(* IEC 61131-3 sources: axsharp/src/ix.compiler/src/Ix.ixc-doc/samples/ax/src, 10 files *)

(* ---- measurement.st ---- *)
NAMESPACE MeasurementExample
    {#ix-attr:[Container(Layout.Wrap)]}
    {#ix-attr:[Group(GroupLayout.GroupBox)]}
    CLASS PUBLIC Measurement
        VAR PUBLIC
            {#ix-set:AttributeName = "Minimum"}
            Min : REAL;
            {#ix-set:AttributeName = "Measured"}
            {#ix-attr:[ReadOnly()]}
            Acquired : REAL;
            {#ix-set:AttributeName = "Maximum"}
            Max : REAL;
            {#ix-set:AttributeName = "Measurement Result"}
            Result : Result;
        END_VAR
    END_CLASS

    TYPE
        Result : INT (
            None := 0,
            Passed := 10,
            Failed := 20
        );
    END_TYPE

    CLASS PUBLIC Measurements
        VAR PUBLIC
            {#ix-attr:[Container(Layout.Stack)]}
            {#ix-attr:[Group(GroupLayout.GroupBox)]}
            {#ix-set:AttributeName = "Stack panel"}
            measurement_stack : Measurement;

            {#ix-attr:[Container(Layout.Wrap)]}
            {#ix-attr:[Group(GroupLayout.GroupBox)]}
            {#ix-set:AttributeName = "Wrap panel"}
            measurement_wrap : Measurement;

            {#ix-attr:[Container(Layout.UniformGrid)]}
            {#ix-attr:[Group(GroupLayout.GroupBox)]}
            {#ix-set:AttributeName = "Grid"}
            measurement_grid : Measurement;

            {#ix-attr:[Container(Layout.Tabs)]}
            {#ix-attr:[Group(GroupLayout.GroupBox)]}
            {#ix-set:AttributeName = "Tabs"}
            measurement_tabs : Measurement;
        END_VAR
    END_CLASS
END_NAMESPACE

(* ---- weather.st ---- *)
{#ix[Container(Layout.Tabs)]}
CLASS weather
    VAR PUBLIC
        GeoLocation : GeoLocation;
        {#ix[Container(Layout.Wrap)]}
        Temperature : REAL;
        Humidity : REAL;
        Location : STRING;
        ChillFactor : REAL;
        Feeling : Feeling;
    END_VAR
END_CLASS

CLASS weathers
    VAR PUBLIC
        i : ARRAY[0..50] OF weatherBase;
    END_VAR
END_CLASS

TYPE
    Feeling : (Freezing, Cold, Lookworm, Warm, Hot);
END_TYPE

TYPE
    Colors : INT (
        RED := 12,
        GREEN := 14,
        BLUE := 23
    );
END_TYPE

(* ---- all_primitives.st ---- *)
CLASS all_primitives
    VAR PUBLIC
        myBOOL	        :       BOOL	      ;
        myBYTE	        :       BYTE	      ;
        myWORD	        :       WORD	      ;
        myDWORD	        :       DWORD	      ;
        myLWORD	        :       LWORD	      ;
        mySINT	        :       SINT	      ;
        myINT	        :       INT	          ;
        myDINT	        :       DINT	      ;
        myLINT	        :       LINT	      ;
        myUSINT	        :       USINT	      ;
        myUINT	        :       UINT	      ;
        myUDINT	        :       UDINT	      ;
        myULINT	        :       ULINT	      ;
        myREAL	        :       REAL	      ;
        myLREAL	        :       LREAL	      ;
        myTIME	        :       TIME	      ;
        myLTIME	        :       LTIME	      ;
        myDATE	        :       DATE	      ;
     //   myLDATE	        :       LDATE	      ;
        myTIME_OF_DAY	:       TIME_OF_DAY	  ;
     //   myLTIME_OF_DAY	:       LTIME_OF_DAY  ;
        myDATE_AND_TIME  :      DATE_AND_TIME ;
     //   myLDATE_AND_TIME :      LDATE_AND_TIME;
     //   myCHAR	        :       CHAR	      ;
     //   myWCHAR	        :       WCHAR	      ;
        mySTRING	        :   STRING	      ;
        myWSTRING	    :       WSTRING	      ;
    END_VAR

END_CLASS

(* ---- example.st ---- *)
CLASS example
    VAR PUBLIC
        {#ix-attr:[Container(Layout.Stack)]}
        primitives_stack: test_primitive;
        {#ix-attr:[Container(Layout.Wrap)]}
        primitives_wrap: test_primitive;
        {#ix-attr:[Container(Layout.Tabs)]}
        primitives_tabs: test_primitive;
        {#ix-attr:[Container(Layout.UniformGrid)]}
        primitives_uniform: test_primitive;

        {#ix-attr:[Container(Layout.Stack)]}
        {#ix-attr:[Group(GroupLayout.GroupBox)]}
        test_groupbox: test_primitive;

        {#ix-attr:[Container(Layout.Stack)]}
        {#ix-attr:[Group(GroupLayout.Border)]}
        test_border: test_primitive;

        {#ix-attr:[Container(Layout.Tabs)]}
        {#ix-attr:[Group(GroupLayout.GroupBox)]}
        testgroupbox: groupbox;
        testborder: border;

        ixcomponent_instance: ixcomponent;
        ixcomponent_instance2: MySecondNamespace.ixcomponent;
        ixcomponent_instance3: ThirdNamespace.ixcomponent;

        refIxComponent : REF_TO ixcomponent;
    END_VAR

    METHOD PUBLIC ReferenceToComponent : Int
        refIxComponent^ := ixcomponent_instance;
    END_METHOD

END_CLASS

(* ---- geolocation.st ---- *)
{#ix-attr:[Container(Layout.Stack)]}
{#ix-attr:[Group(GroupLayout.GroupBox)]}
{#ix-set:AttributeName = "Location"}
CLASS  GeoLocation
    VAR PUBLIC
        {#ix-set:AttributeName = "Latitude [°]"}
        {#ix-set:AttributeMinimum = -90.0f}
        {#ix-set:AttributeMaximum = 90.0f}
        Latitude : REAL;
        {#ix-set:AttributeName = "Logitude [°]"}
        {#ix-set:AttributeMinimum = 0.0f}
        {#ix-set:AttributeMaximum = 180.0f}
        Longitude : REAL;
        {#ix-set:AttributeName = "Altitude [m]"}
        Altitude : REAL;
        {#ix-set:AttributeName = "Short descriptor"}
        Description : STRING[10];
        {#ix-set:AttributeName = "Long descriptor"}
        LongDescription : STRING[254];
    END_VAR
END_CLASS

(* ---- ixcomponent.st ---- *)
CLASS ixcomponent
    VAR PUBLIC
        {#ix-set:AttributeName = "My integer"}
        my_int : INT;
        {#ix-set:AttributeName = "My string"}
        my_string : STRING;
        {#ix-set:AttributeName = "My bool"}
        my_bool : BOOL;
    END_VAR
END_CLASS

NAMESPACE MySecondNamespace
    CLASS ixcomponent
        VAR PUBLIC
            {#ix-set:AttributeName = "My integer"}
            my_int : INT;
            {#ix-set:AttributeName = "My string"}
            my_string : STRING;
            {#ix-set:AttributeName = "My bool"}
            my_bool : BOOL;
        END_VAR
    END_CLASS
END_NAMESPACE

NAMESPACE ThirdNamespace
    CLASS ixcomponent
        VAR PUBLIC
            {#ix-set:AttributeName = "My integer"}
            my_int : INT;
            {#ix-set:AttributeName = "My string"}
            my_string : STRING;
            {#ix-set:AttributeName = "My bool"}
            my_bool : BOOL;
        END_VAR
    END_CLASS
END_NAMESPACE

(* ---- monster.st ---- *)
NAMESPACE MonsterData
    CLASS MonsterBase
        VAR PUBLIC
            ArrayOfBytes : ARRAY[0..3] OF BYTE;
            ArrayOfDrives : ARRAY[0..3] OF DriveBase;
            ArrayOfIxComponent : ARRAY[0..3] OF ixcomponent;
        END_VAR
    END_CLASS
    CLASS Monster EXTENDS MonsterBase
        VAR PUBLIC
            DriveA : DriveBase;
        END_VAR
    END_CLASS

    CLASS DriveBase
        VAR PUBLIC
            Position : LREAL;
            Velo : LREAL;
            Acc : LREAL;
            Dcc : LREAL;
        END_VAR
    END_CLASS
END_NAMESPACE

(* ---- weatherBase.st ---- *)
    {#ix-attr:[Container(Layout.Stack)]}
    {#ix-attr:[Group(GroupLayout.GroupBox)]}
    CLASS PUBLIC weatherBase
      VAR PUBLIC
        Latitude : REAL;
        Longitude : REAL;
        Altitude : REAL;
        Description : STRING;
        {#ix-attr:[ReadOnly()]}
        LongDescription : STRING;
        {#ix-attr:[ReadOnce()]}
        {#ix-set:AttributeName = "this has [ReadOnce()] attribute will be readon only once..."}
        StartCounter : INT;

        {#ix-attr:[RenderIgnore()]}
        {#ix-set:AttributeName = "[RenderIgnore()] must not be displayed!"}
        RenderIgnoreAllToghether : STRING;
        {#ix-set:AttributeName = "[RenderIgnore(''Control'')]"}
        {#ix-attr:[RenderIgnore("Control")]}
        RenderIgnoreWhenControl : STRING;
        {#ix-set:AttributeName = "[RenderIgnore(''Display'')]"}
        {#ix-attr:[RenderIgnore("Display")]}
        RenderIgnoreWhenDisplay : STRING;
        {#ix-set:AttributeName = "[RenderIgnore(''Control'', ''ShadowControl'')]"}
        {#ix-attr:[RenderIgnore("Control", "ShadowControl")]}
        RenderIgnoreWhenControlAndShadow : STRING;
        {#ix-set:AttributeName = "[RenderIgnore(''Display'', ''ShadowDisplay'')]"}
        {#ix-attr:[RenderIgnore("Display", "ShadowDisplay")]}
        RenderIgnoreWhenDisplayAndShadow : STRING;
      END_VAR
    END_CLASS

(* ---- configuration.st ---- *)
USING MonsterData;
CONFIGURATION MyConfiguration
    TASK Main(Interval := T#10ms, Priority := 1);
    PROGRAM P1 WITH Main: MyProgram;

    VAR_GLOBAL
        all_primitives : all_primitives;
        weather : weather;
        weathers : weathers;
        {#ix-set:AttributeName = "Weather in a stack pannel and grouped in group box"}
        weather_stacked : Layouts.Stacked.weather;
        {#ix-set:AttributeName = "Weather in a wrap pannel and grouped in group box"}
        weather_wrapped : Layouts.Wrapped.weather;
        {#ix-set:AttributeName = "Weather in a tabs and grouped in group box"}
        weather_tabbed : Layouts.Tabbed.weather;
        {#ix-set:AttributeName = "Weather structure set to read once"}
        {#ix-attr:[ReadOnce()]}
        weather_readOnce : Layouts.Stacked.weather;
        {#ix-set:AttributeName = "Weather structure set to read only"}
        {#ix-attr:[ReadOnly()]}
        weather_readOnly : Layouts.Stacked.weather;

        test_example: example;
        measurements : MeasurementExample.Measurements;
        monster : Monster;
    END_VAR
END_CONFIGURATION

(* ---- program.st ---- *)
PROGRAM MyProgram
    VAR_EXTERNAL
        all_primitives : all_primitives;
        weather_stacked : Layouts.Stacked.weather;
        weather_wrapped : Layouts.Wrapped.weather;
        weather_tabbed : Layouts.Tabbed.weather;
        weather_readOnce : Layouts.Stacked.weather;
        test_example: example;
    END_VAR

    VAR

    END_VAR

    VAR_TEMP

    END_VAR
    all_primitives.myINT := all_primitives.myINT + 1;
    weather_stacked.Altitude := all_primitives.myINT;
    weather_wrapped.Altitude := all_primitives.myINT;
    weather_tabbed.Altitude := all_primitives.myINT;
    weather_readOnce.Altitude := all_primitives.myINT;

    weather_stacked.StartCounter := all_primitives.myINT;
    weather_wrapped.StartCounter := all_primitives.myINT;
    weather_tabbed.StartCounter := all_primitives.myINT;
    weather_readOnce.StartCounter := all_primitives.myINT;

    test_example.ReferenceToComponent();

END_PROGRAM
